Fanuc KAREL source: kb00106.KL

PROGRAM KB00106
%STACKSIZE=65535
%PRIORITY=65535
%NOLOCKGROUP
-- UNRESOLVED DECLARATIONS (source type spelling not recovered)
-- P1 : TYPE_0x1100 (type_u16=0x1100)
BEGIN
INIT_QUEUE(P1)
END KB00106
